ABB RobotStudio station: ABB_IRB_1300.rsstnx

Station ABB_IRB_1300_Neu_1 (saved by RobotStudio 26.2.11700.0)
Controller Steuerung_ABB_IRB_1300, task T_ROB1: task frame (RAPID world) sits at (0, 0, 775) mm, rotated rx 0 ry 0 rz 30 deg in the station
Controller Steuerung_ABB_IRB_1300
  mechanical unit ROB_1: Roboter_ABB_IRB_1300, 6 joints, base frame (0, 0, 0) mm
Layout (positions relative to the parent item):
  - Roboter_ABB_IRB_1300 [mechanism, from %ABB.RobotStudio.Models.IRB1300%\IRB1300_7_140__01.rslib] at (0, 0, 775) mm, rotated rx 0 ry 0 rz 30 deg; joint values [-0.5236, -0.9812, 0.8606, 0, 0.6441, 0] (rad or m)
  - Keyence_Modul1 [graphiccomponentgroup] at (856, 0, 1037) mm, rotated rx 0 ry 0 rz 90 deg
    - DEFAULT [part] at (0, -2, 57.1) mm, size 122.5 x 88.9 x 126.5 mm
    - DEFAULT [part] at (0, -73.1, 67.5) mm, size 145.3 x 131.6 x 127.1 mm
    - DEFAULT [part] at (0, -127.8, 26) mm, size 184.3 x 146.8 x 135.3 mm
    - DEFAULT [part] at (59.9, -20, 61.2) mm, rotated rx 0 ry 90 rz 0 deg, size 61.9 x 49.3 x 15.5 mm
    - DEFAULT [part] at (-59.9, -20, 10) mm, rotated rx 0 ry -90 rz 0 deg, size 52 x 39 x 15.4 mm
  - Keyence_Modul4 [graphiccomponentgroup] at (-856, 0, 1037) mm, rotated rx 0 ry 0 rz -90 deg
    - DEFAULT [part] at (0, -2, 57.1) mm, size 120 x 86.2 x 124.5 mm
    - DEFAULT [part] at (0, -73.1, 67.5) mm, size 143 x 130 x 125 mm
    - DEFAULT [part] at (0, -127.8, 26) mm, size 181.4 x 145 x 132.1 mm
    - DEFAULT [part] at (59.9, -20, 61.2) mm, rotated rx 0 ry 90 rz 0 deg, size 60.9 x 48.3 x 14.6 mm
    - DEFAULT [part] at (-59.9, -20, 10) mm, rotated rx 0 ry -90 rz 0 deg, size 51.2 x 38.5 x 14.9 mm
  - Keyence_Modul6 [graphiccomponentgroup] at (428, 741.32, 1037) mm, rotated rx 0 ry 0 rz 150 deg
    - DEFAULT [part] at (0, -2, 57.1) mm, size 120 x 86.2 x 124.5 mm
    - DEFAULT [part] at (0, -73.1, 67.5) mm, size 143 x 130 x 125 mm
    - DEFAULT [part] at (0, -127.8, 26) mm, size 181.4 x 145 x 132.1 mm
    - DEFAULT [part] at (59.9, -20, 61.2) mm, rotated rx 0 ry 90 rz 0 deg, size 60.9 x 48.3 x 14.6 mm
    - DEFAULT [part] at (-59.9, -20, 10) mm, rotated rx 0 ry -90 rz 0 deg, size 51.2 x 38.5 x 14.9 mm
  - Keyence_Modul3 [graphiccomponentgroup] at (-428, -741.32, 1037) mm, rotated rx 0 ry 0 rz -30 deg
    - DEFAULT [part] at (0, -2, 57.1) mm, size 120 x 86.2 x 124.5 mm
    - DEFAULT [part] at (0, -73.1, 67.5) mm, size 143 x 130 x 125 mm
    - DEFAULT [part] at (0, -127.8, 26) mm, size 181.4 x 145 x 132.1 mm
    - DEFAULT [part] at (59.9, -20, 61.2) mm, rotated rx 0 ry 90 rz 0 deg, size 60.9 x 48.3 x 14.6 mm
    - DEFAULT [part] at (-59.9, -20, 10) mm, rotated rx 0 ry -90 rz 0 deg, size 51.2 x 38.5 x 14.9 mm
  - Keyence_Modul5 [graphiccomponentgroup] at (-428, 741.32, 1037) mm, rotated rx 0 ry 0 rz -150 deg
    - DEFAULT [part] at (0, -2, 57.1) mm, size 120 x 86.2 x 124.5 mm
    - DEFAULT [part] at (0, -73.1, 67.5) mm, size 143 x 130 x 125 mm
    - DEFAULT [part] at (0, -127.8, 26) mm, size 181.4 x 145 x 132.1 mm
    - DEFAULT [part] at (59.9, -20, 61.2) mm, rotated rx 0 ry 90 rz 0 deg, size 60.9 x 48.3 x 14.6 mm
    - DEFAULT [part] at (-59.9, -20, 10) mm, rotated rx 0 ry -90 rz 0 deg, size 51.2 x 38.5 x 14.9 mm
  - Keyence_Modul2 [graphiccomponentgroup] at (428, -741.32, 1037) mm, rotated rx 0 ry 0 rz 30 deg
    - DEFAULT [part] at (0, -2, 57.1) mm, size 120 x 86.2 x 124.5 mm
    - DEFAULT [part] at (0, -73.1, 67.5) mm, size 143 x 130 x 125 mm
    - DEFAULT [part] at (0, -127.8, 26) mm, size 181.4 x 145 x 132.1 mm
    - DEFAULT [part] at (59.9, -20, 61.2) mm, rotated rx 0 ry 90 rz 0 deg, size 60.9 x 48.3 x 14.6 mm
    - DEFAULT [part] at (-59.9, -20, 10) mm, rotated rx 0 ry -90 rz 0 deg, size 51.2 x 38.5 x 14.9 mm
  - Arbeitsplatte [part] at (0, 0, 992) mm, size 1950 x 2230 x 1035 mm
  - Käfig_Modul1 [part] at (1520, 0, 0) mm, size 1090 x 1090 x 2007 mm
  - Käfig_Modul4 [part] at (-1520, 0, 0) mm, size 1090 x 1090 x 2007 mm
  - Käfig_Modul5 [part] at (-760, 1316.36, 0) mm, rotated rx 0 ry 0 rz -60 deg, size 1090 x 1090 x 2007 mm
  - Käfig_Modul2 [part] at (760, -1316.36, 0) mm, rotated rx 0 ry 0 rz -60 deg, size 1090 x 1090 x 2007 mm
  - Käfig_Modul3 [part] at (-760, -1316.36, 0) mm, rotated rx 0 ry 0 rz 60 deg, size 1090 x 1090 x 2007 mm
  - Käfig_Modul6 [part] at (760, 1316.36, 0) mm, rotated rx 0 ry 0 rz 60 deg, size 1090 x 1090 x 2007 mm
Targets, tools, work objects and paths stored in the station, written as RAPID:
! task T_ROB1
MODULE CalibData
  PERS wobjdata coordinate_system_module_5:=[FALSE,TRUE,"",[[-499.960321416,1020.013088225,257.5],[1,0,0,0.000005866]],[[0,0,0],[1,0,0,0]]];
  PERS wobjdata coordinate_system_module_2:=[FALSE,TRUE,"",[[498.985385611,-1020.52304872,257.5],[0.000473151,0,0,-0.999999888]],[[0,0,0],[1,0,0,0]]];
  PERS wobjdata coordinate_system_module_1:=[FALSE,TRUE,"",[[1134.907540478,-83.031342842,257.5],[0.500647833,0,0,-0.865651054]],[[0,0,0],[1,0,0,0]]];
  PERS wobjdata coordinate_system_module_3:=[FALSE,TRUE,"",[[-636.650058157,-941.997300822,257.5],[0.50036151,0,0,0.865816585]],[[0,0,0],[1,0,0,0]]];
  PERS wobjdata coordinate_system_module_4:=[FALSE,TRUE,"",[[-1133.976818569,78.784535634,257.5],[0.86565239,0,0,0.500645524]],[[0,0,0],[1,0,0,0]]];
  PERS wobjdata coordinate_system_module_6:=[FALSE,TRUE,"",[[638.159114859,940.449669808,257.5],[0.866179246,-0,0,-0.499733442]],[[0,0,0],[1,0,0,0]]];
ENDMODULE

